Staubli VAL3: movePoint.pgx

program movePoint(num x_nIndex)
  local bool l_bResult
  local jointRx l_joint
begin
  l_bResult=userPageConfirm("是否移动到点位："+toString("",x_nIndex)+"?")
  if l_bResult and rs:_nOmacStat==9
    resetMotion()
    l_bResult=pointToJoint(flange,herej(),safeTemp:sSPoint[x_nIndex].pPointRx,l_joint)
    if l_bResult
      movej(safeTemp:sSPoint[x_nIndex].pPointRx,flange,mSimulate)
    else
      popUpMsg("无法移动到该安全点位")
    endIf
  endIf
  if rs:_nOmacStat!=9
    userPageAlert("机器人当前状态不满足，无法执行移动")
  endIf
end
